SUBAPPLICATION Uebung_154 (* Stoßfreie Hand/Auto-Umschaltung CTRL_PID_AR, simulierte PT1-Strecke *)
  (* Standard: 61499-2; Description: Copyright (c) 2026 Meisterschulen am Ostbahnhof This program and the accompanying materials are made available under the terms of the Eclipse Public License 2.0 which is available at https://www.eclipse.org/legal/epl-2.0/ SPDX-License-Identifier: EPL-2.0 *)
  (* Version 1.0, 2026-11-15, Franz Höpfinger, Meisterschulen am Ostbahnhof, initial API and implementation and/or initial documentation *)
  PACKAGE Uebungen;
  IMPORT logiBUS::io::DI::logiBUS_DI::Input_I1;
  IMPORT logiBUS::io::DI::logiBUS_DI::Input_I2;
  IMPORT logiBUS::io::DI::logiBUS_DI::Input_I3;
  IMPORT logiBUS::io::DI::logiBUS_DI_Events::BUTTON_SINGLE_CLICK;
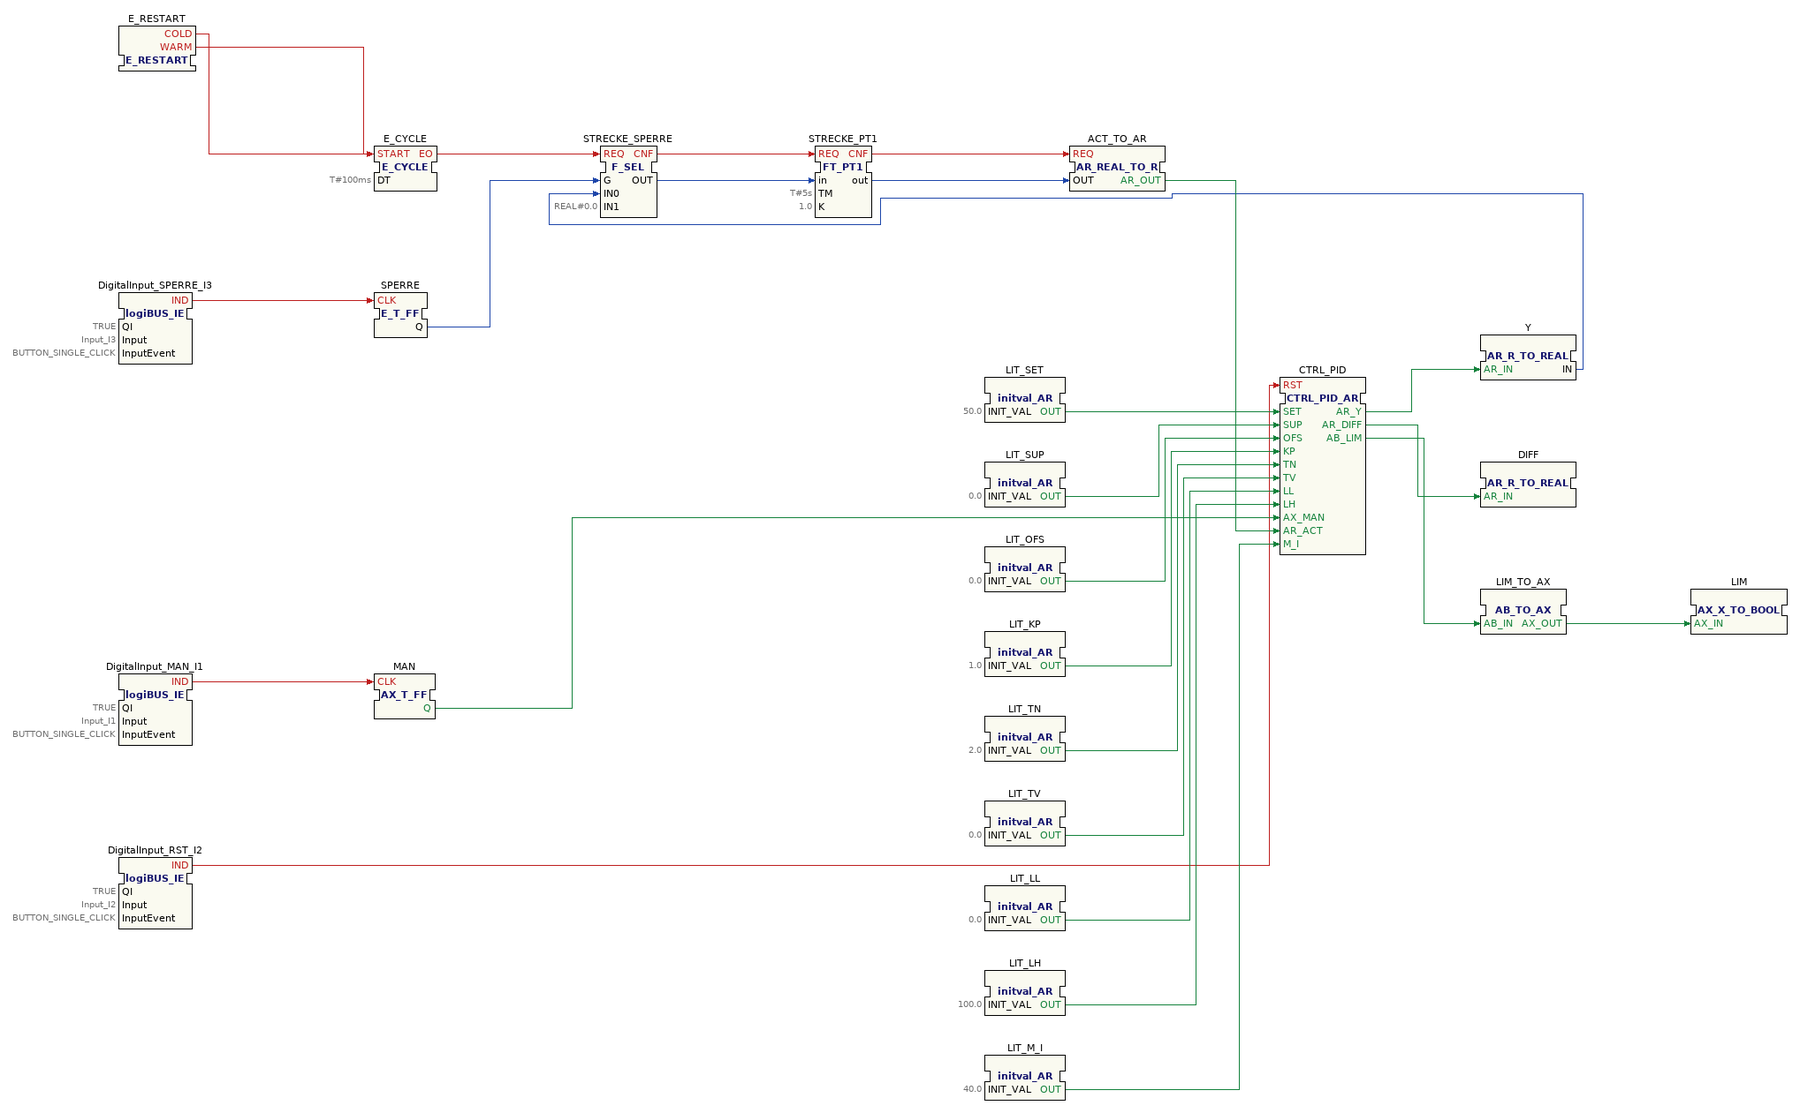
  (* Test stoßfreie Hand/Auto-Umschaltung (CTRL_PID_AR, OSCAT-Fix #385) Strecke simuliert: PT1 (5 s) aus Y, Takt 100 ms, startet von selbst. I1 = Hand/Auto (Start: Auto), I2 = RST Integrator, I3 = Ausgang sperren (Strecke bekommt 0). Handwert M_I: 40 (fest, LIT_M_I). Watch: Y.IN, STRECKE_PT1.out (Istwert), DIFF.IN, LIM.IN. 1) I1 Hand: Y = M_I. I1 Auto: Y springt nicht, regelt von M_I aus weiter. 2) Start in Auto: Y beginnt bei 50 (KP*DIFF), läuft nicht erst bis LH hoch. 3) Gegenprobe: in Auto I2 drücken -> Integrator 0, Y springt auf KP*DIFF. 4) Windup: I3 sperren -> Istwert fällt, Y läuft bis LH (100), LIM = TRUE. Lösung im Projekt: RST bei steigender Freigabe. *)
  FBS
    CTRL_PID : OSCAT_adapter::Control::CTRL_PID_AR;
    LIT_SET : adapter::types::unidirectional::AR::initval::initval_AR(INIT_VAL := 50.0);
    LIT_SUP : adapter::types::unidirectional::AR::initval::initval_AR(INIT_VAL := 0.0);
    LIT_OFS : adapter::types::unidirectional::AR::initval::initval_AR(INIT_VAL := 0.0);
    LIT_KP : adapter::types::unidirectional::AR::initval::initval_AR(INIT_VAL := 1.0);
    LIT_TN : adapter::types::unidirectional::AR::initval::initval_AR(INIT_VAL := 2.0);
    LIT_TV : adapter::types::unidirectional::AR::initval::initval_AR(INIT_VAL := 0.0);
    LIT_LL : adapter::types::unidirectional::AR::initval::initval_AR(INIT_VAL := 0.0);
    LIT_LH : adapter::types::unidirectional::AR::initval::initval_AR(INIT_VAL := 100.0);
    E_RESTART : iec61499::events::E_RESTART;
    SPERRE : iec61499::events::E_T_FF;
    MAN : adapter::events::unidirectional::AX_T_FF;
    Y : adapter::conversion::unidirectional::AR_R_TO_REAL;
    DIFF : adapter::conversion::unidirectional::AR_R_TO_REAL;
    LIM_TO_AX : adapter::conversion::unidirectional::AB_TO_AX;
    LIM : adapter::conversion::unidirectional::AX_X_TO_BOOL;
    DigitalInput_MAN_I1 : logiBUS::io::DI::logiBUS_IE(QI := TRUE, Input := Input_I1, InputEvent := BUTTON_SINGLE_CLICK);
    DigitalInput_RST_I2 : logiBUS::io::DI::logiBUS_IE(QI := TRUE, Input := Input_I2, InputEvent := BUTTON_SINGLE_CLICK);
    DigitalInput_SPERRE_I3 : logiBUS::io::DI::logiBUS_IE(QI := TRUE, Input := Input_I3, InputEvent := BUTTON_SINGLE_CLICK);
    E_CYCLE : iec61499::events::E_CYCLE(DT := T#100ms);
    STRECKE_SPERRE : iec61131::selection::F_SEL(IN1 := REAL#0.0);
    STRECKE_PT1 : OSCAT::Basic::POUs::Engineering::Control::FT_PT1(TM := T#5s, K := 1.0);
    ACT_TO_AR : adapter::conversion::unidirectional::AR_REAL_TO_R;
    LIT_M_I : adapter::types::unidirectional::AR::initval::initval_AR(INIT_VAL := 40.0);
  END_FBS
  EVENT_CONNECTIONS
    E_RESTART.COLD TO E_CYCLE.START;
    E_RESTART.WARM TO E_CYCLE.START;
    E_CYCLE.EO TO STRECKE_SPERRE.REQ;
    STRECKE_SPERRE.CNF TO STRECKE_PT1.REQ;
    STRECKE_PT1.CNF TO ACT_TO_AR.REQ;
    DigitalInput_SPERRE_I3.IND TO SPERRE.CLK;
    DigitalInput_MAN_I1.IND TO MAN.CLK;
    DigitalInput_RST_I2.IND TO CTRL_PID.RST;
  END_CONNECTIONS
  DATA_CONNECTIONS
    SPERRE.Q TO STRECKE_SPERRE.G;
    Y.IN TO STRECKE_SPERRE.IN0;
    STRECKE_SPERRE.OUT TO STRECKE_PT1.in;
    STRECKE_PT1.out TO ACT_TO_AR.OUT;
  END_CONNECTIONS
  ADAPTER_CONNECTIONS
    LIT_SET.OUT TO CTRL_PID.SET;
    LIT_SUP.OUT TO CTRL_PID.SUP;
    LIT_OFS.OUT TO CTRL_PID.OFS;
    LIT_KP.OUT TO CTRL_PID.KP;
    LIT_TN.OUT TO CTRL_PID.TN;
    LIT_TV.OUT TO CTRL_PID.TV;
    LIT_LL.OUT TO CTRL_PID.LL;
    LIT_LH.OUT TO CTRL_PID.LH;
    MAN.Q TO CTRL_PID.AX_MAN;
    CTRL_PID.AR_Y TO Y.AR_IN;
    CTRL_PID.AR_DIFF TO DIFF.AR_IN;
    CTRL_PID.AB_LIM TO LIM_TO_AX.AB_IN;
    LIM_TO_AX.AX_OUT TO LIM.AX_IN;
    ACT_TO_AR.AR_OUT TO CTRL_PID.AR_ACT;
    LIT_M_I.OUT TO CTRL_PID.M_I;
  END_CONNECTIONS
END_SUBAPPLICATION
